// TIA Portal V20 export
// export: Created 2026-10-12T05:42:34.3523902Z, ExportSetting WithDefaults, DisplayName Totally Integrated Automation Portal, DisplayVersion V20, DisplayName TIA Portal Openness, DisplayVersion V20, DisplayName TIA Portal Teamcenter Gateway, DisplayVersion V20, DisplayName TIA Portal Version Control Interface, DisplayVersion V20, DisplayName SINAMICS Startdrive Advanced, DisplayVersion V20 SP1 Update 2, DisplayName SINAMICS Startdrive G110M, G120, G120C, G120D, G120P, G115D, DisplayVersion V20 SP1 Update 2, DisplayName SINAMICS Startdrive G130, G150, S120, S150, SINAMICS MV, G220, S200, S210, DisplayVersion V20 SP1 Update 2, DisplayName STEP 7 Professional, DisplayVersion V20, DisplayName STEP 7 Safety, DisplayVersion V20, DisplayName WinCC Basic/Comfort/Advanced, DisplayVersion V20, DisplayName WinCC Professional, DisplayVersion V20, DisplayName WinCC Unified, DisplayVersion V20
FUNCTION "F_PressDemoDoorClose" : Void   // FC162, SCL
{ S7_Optimized_Access := 'TRUE' }
VERSION : 0.1
// stored: AutoNumber true, IsIECCheckEnabled false, SetENOAutomatically false, UDAEnableTagReadback false
   VAR_INPUT
      Closed : Bool;
      TwoHandHeld : Bool;
      RequireTwoHandStart : Bool;
      SourcePath : String;
   END_VAR
   VAR_IN_OUT
      Seq : "FRK_SequenceCtx";
      AlarmLog : "FRK_AlarmLog";
   END_VAR
   VAR_TEMP
      Held : Bool;
      Diag : "ST_Diagnostic";
   END_VAR
BEGIN

   #Held := "FRK_SeqAwait"(Seq := #Seq, Label := 'project.condition.twoHandHeldDuringDoorClose', Ok := #TwoHandHeld OR NOT #RequireTwoHandStart);
   "FRK_SeqSelect"(Seq := #Seq,
                   AdvanceOk := #Closed,
                   Jump1Ok := NOT #Held);
   IF #Seq.RetVal = 2 THEN
       #Diag := "FRK_UnitScratch".EmptyDiagnostic;
       #Diag.ReasonCode := 12001;
       #Diag.Description := WSTRING#'project.warning.twoHandReleasedDuringDoorClose';
       #Diag.SourcePath := STRING_TO_WSTRING(#SourcePath);
       #Diag.Severity := 0;
       #Diag.Category := 0;
       "FRK_SeqMessage"(Seq := #Seq,
                        AlarmLog := #AlarmLog,
                        Diag := #Diag);
   END_IF;
END_FUNCTION
